// TIA Portal V21 program export: 3 tag tables, 0 data types, 5 data blocks, 7 code blocks (in call order from the OBs), 0 instance data blocks

VAR_GLOBAL   // PLC tag table "DI"
   "DI_PRODUCT SENSOR" AT %I0.0 : Bool;
   "DI_AUTO MANUAL SELECTION" AT %I0.1 : Bool;
   "DI_CYCLE START PB" AT %I0.2 : Bool;
   "DI_CYCLE STOP PB" AT %I0.3 : Bool;
   "DI_EMERGENCY PB" AT %I0.4 : Bool;
   "DI_CONVEYOR VFD FAULT" AT %I0.5 : Bool;
   "DI_SPARE I0.6" AT %I0.6 : Bool;
   "DI_SPARE I0.7" AT %I0.7 : Bool;
   "DI_SPARE I1.0" AT %I1.0 : Bool;
   "DI_SPARE I1.1" AT %I1.1 : Bool;
   "DI_SPARE I1.2" AT %I1.2 : Bool;
   "DI_SPARE I1.3" AT %I1.3 : Bool;
   "DI_SPARE I1.4" AT %I1.4 : Bool;
   "DI_SPARE I1.5" AT %I1.5 : Bool;
END_VAR

VAR_GLOBAL   // PLC tag table "DO"
   "DO_CONVEYOR FWD ON" AT %Q0.0 : Bool;
   "DO_CONVEYOR REV ON" AT %Q0.1 : Bool;
   "DO_FAULT RESET" AT %Q0.2 : Bool;
   "DO_TL GREEN" AT %Q0.3 : Bool;
   "DO_TL RED" AT %Q0.4 : Bool;
   "DO_TL AMBER" AT %Q0.5 : Bool;
   "DO_SPARE Q0.6" AT %Q0.6 : Bool;
   "DO_SPARE Q0.7" AT %Q0.7 : Bool;
   "DO_SPARE Q1.0" AT %Q1.0 : Bool;
   "DO_SPARE Q1.1" AT %Q1.1 : Bool;
END_VAR

VAR_GLOBAL   // PLC tag table "Default tag table"
   System_Byte AT %MB1 : Byte;
   FirstScan AT %M1.0 : Bool;
   DiagStatusUpdate AT %M1.1 : Bool;
   AlwaysTRUE AT %M1.2 : Bool;
   AlwaysFALSE AT %M1.3 : Bool;
   Clock_Byte AT %MB0 : Byte;
   Clock_10Hz AT %M0.0 : Bool;
   Clock_5Hz AT %M0.1 : Bool;
   "Clock_2.5Hz" AT %M0.2 : Bool;
   Clock_2Hz AT %M0.3 : Bool;
   "Clock_1.25Hz" AT %M0.4 : Bool;
   Clock_1Hz AT %M0.5 : Bool;
   "Clock_0.625Hz" AT %M0.6 : Bool;
   "Clock_0.5Hz" AT %M0.7 : Bool;
   "CONTROL ON FLAG" AT %M2.0 : Bool;
   "MANUAL MODE SELECTED" AT %M2.1 : Bool;
   "AUTO MODE SELECTED" AT %M2.2 : Bool;
   "FAULT RESET FLAG" AT %M2.3 : Bool;
   "FAULT BIT" AT %M2.4 : Bool;
   "MANUAL CONVEYOR FWD ON FLAG" AT %M2.5 : Bool;
   "MANUAL CONVEYOR REV ON FLAG" AT %M2.6 : Bool;
END_VAR

DATA_BLOCK "DB_ALARMS"   // DB2
{ S7_Optimized_Access := 'FALSE' }
VERSION : 0.1
// stored: AutoNumber true, DBAccessibleFromOPCUA true, IsOnlyStoredInLoadMemory false, IsWriteProtectedInAS false
   VAR
      "EMERGENCY PB PRESSED FAULT" : Bool;
      "VFD FAULT" : Bool;
      SPARE1 : Bool;
      SPARE2 : Bool;
      SPARE3 : Bool;
      SPARE4 : Bool;
      SPARE5 : Bool;
      SPARE6 : Bool;
      SPARE7 : Bool;
      SPARE8 : Bool;
      SPARE9 : Bool;
      SPARE10 : Bool;
      SPARE11 : Bool;
      SPARE12 : Bool;
      SPARE13 : Bool;
      SPARE14 : Bool;
      "FAULT POP" : Bool;
      "WARNING POP" : Bool;
   END_VAR
BEGIN
END_DATA_BLOCK

DATA_BLOCK "DB_AUTO"   // DB3
{ S7_Optimized_Access := 'FALSE' }
VERSION : 0.1
// stored: AutoNumber true, DBAccessibleFromOPCUA true, IsOnlyStoredInLoadMemory false, IsWriteProtectedInAS false
   VAR
      ACTIVE : Bool;
      "CONVEYOR ON" : Bool;
      "CONVEYOR OFF1" : Bool;
      "CONVEYOR OFF2" : Bool;
      P_TRG : Bool;
      "CAMERA DONE" : Bool;
      "AUTO STATUS" : Int;
      "STOP DELAY TIMER" : IEC_TIMER;
      "SENSOR CHECK DELAY" { S7_SetPoint := 'True'} : IEC_TIMER;
   END_VAR
BEGIN
END_DATA_BLOCK

DATA_BLOCK "DB_CAMERA"   // DB5
{ S7_Optimized_Access := 'FALSE' }
VERSION : 0.1
// stored: AutoNumber true, DBAccessibleFromOPCUA true, IsOnlyStoredInLoadMemory false, IsWriteProtectedInAS false
   VAR
      DATA1 : Int;
      DATA2 : Int;
      DATA3 : Int;
      DATA4 : Int;
      DATA5 : Int;
      DATA6 : Int;
      DATA7 : Int;
      DATA8 : Int;
      DATA9 : Int;
      DATA10 : Int;
      DATA11 : Int;
      DATA12 : Int;
      DATA13 : Int;
      DATA14 : Int;
      DATA15 : Int;
      DATA16 : Int;
      DATA17 : Int;
      DATA18 : Int;
      DATA19 : Int;
   END_VAR
BEGIN
END_DATA_BLOCK

DATA_BLOCK "DB_HMI"   // DB1
{ S7_Optimized_Access := 'FALSE' }
VERSION : 0.1
// stored: AutoNumber true, DBAccessibleFromOPCUA true, IsOnlyStoredInLoadMemory false, IsWriteProtectedInAS false
   VAR RETAIN
      "FAULT RESET PB" : Bool;
      "MOTOR JOG FWD PB" : Bool;
      "MOTOR JOG REV PB" : Bool;
      "STOP TIME" : DInt;
      "CAMERA DONE" : Bool;
   END_VAR
BEGIN
END_DATA_BLOCK

DATA_BLOCK "DB_TCP_IP"   // DB12
{ S7_Optimized_Access := 'TRUE' }
VERSION : 0.1
// stored: AutoNumber true, DBAccessibleFromOPCUA true, IsOnlyStoredInLoadMemory false, IsRetainMemResEnabled false, IsWriteProtectedInAS false, MemoryReserve 100
   VAR
      "MY CONNECT DATA" { S7_SetPoint := 'True'} : TCON_IP_v4;
      "NO OF DONE" { S7_SetPoint := 'True'} : UDInt;
      "NO OF ERROR" : UDInt;
      "ERROR STATUS" : UDInt;
   END_VAR
BEGIN
END_DATA_BLOCK

ORGANIZATION_BLOCK "Main"   // OB1, LAD, ProgramCycle
TITLE = "Main Program Sweep (Cycle)"
{ S7_Optimized_Access := 'TRUE' }
VERSION : 0.1
// stored: AutoNumber true, IsIECCheckEnabled false, SetENOAutomatically false
   VAR_INPUT
      Initial_Call : Bool;   // Initial call of this OB
      Remanence : Bool;   // =True, if remanent data are available
   END_VAR
BEGIN

REGION Network 1
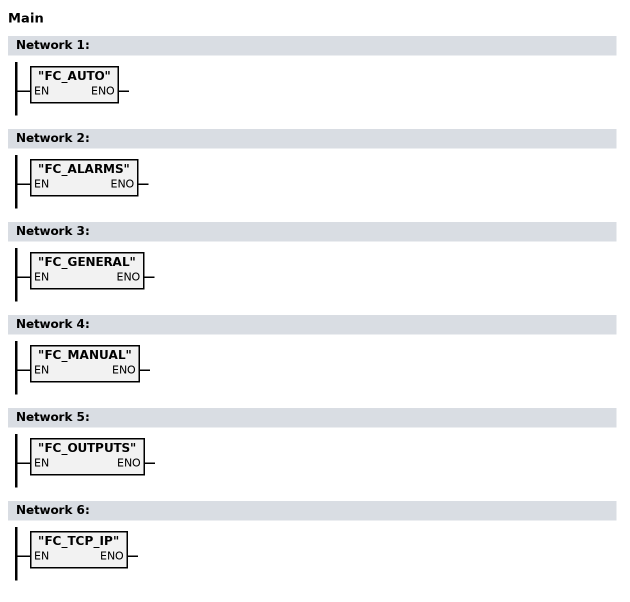
   RUNG wire#powerrail
      "FC_AUTO"()
   END_RUNG
   // the same network as SCL:
   "FC_AUTO"();
END_REGION

REGION Network 2
   RUNG wire#powerrail
      "FC_ALARMS"()
   END_RUNG
   // the same network as SCL:
   "FC_ALARMS"();
END_REGION

REGION Network 3
   RUNG wire#powerrail
      "FC_GENERAL"()
   END_RUNG
   // the same network as SCL:
   "FC_GENERAL"();
END_REGION

REGION Network 4
   RUNG wire#powerrail
      "FC_MANUAL"()
   END_RUNG
   // the same network as SCL:
   "FC_MANUAL"();
END_REGION

REGION Network 5
   RUNG wire#powerrail
      "FC_OUTPUTS"()
   END_RUNG
   // the same network as SCL:
   "FC_OUTPUTS"();
END_REGION

REGION Network 6
   RUNG wire#powerrail
      "FC_TCP_IP"()
   END_RUNG
   // the same network as SCL:
   "FC_TCP_IP"();
END_REGION
END_ORGANIZATION_BLOCK

FUNCTION "FC_AUTO" : Void   // FC5, LAD
{ S7_Optimized_Access := 'TRUE' }
VERSION : 0.1
// stored: AutoNumber true, IsIECCheckEnabled false, SetENOAutomatically false, UDAEnableTagReadback false
   VAR_TEMP   // added for the SCL form of the ladder/FBD networks
      _w1 : Bool;
      _w2 : Bool;
      _w3 : Bool;
   END_VAR
BEGIN

REGION Network 1: AUTO ON
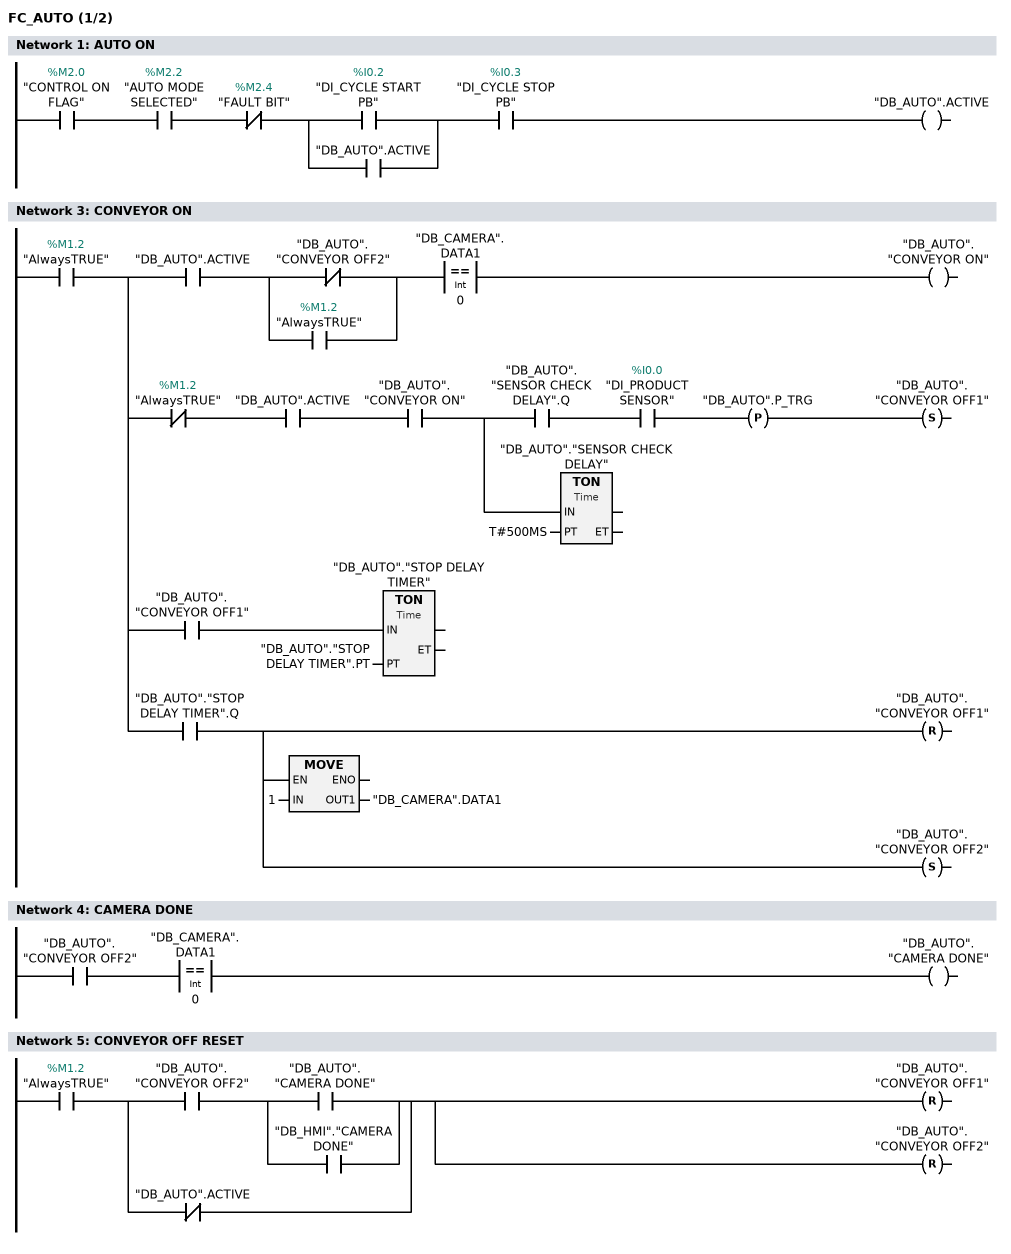
   RUNG wire#powerrail
      Contact( "CONTROL ON FLAG" )
      Contact( "AUTO MODE SELECTED" )
      I_Contact( "FAULT BIT" )
      wire#w1
      Contact( "DI_CYCLE START PB" )
      wire#w2
      Contact( "DI_CYCLE STOP PB" )
      Coil( "DB_AUTO".ACTIVE )
   END_RUNG
   RUNG wire#w1
      Contact( "DB_AUTO".ACTIVE )
   END_RUNG wire#w2
   // the same network as SCL:
   "DB_AUTO".ACTIVE := "CONTROL ON FLAG" AND "AUTO MODE SELECTED" AND NOT "FAULT BIT" AND ("DI_CYCLE START PB" OR "DB_AUTO".ACTIVE) AND "DI_CYCLE STOP PB";
END_REGION

REGION Network 2 (SCL): STOP DELAY TIME
   "DB_AUTO"."STOP DELAY TIMER".PT := "DB_HMI"."STOP TIME" * 1000;
END_REGION

REGION Network 3: CONVEYOR ON
   RUNG wire#powerrail
      Contact( "AlwaysTRUE" )
      wire#w1
      Contact( "DB_AUTO".ACTIVE )
      wire#w2
      I_Contact( "DB_AUTO"."CONVEYOR OFF2" )
      wire#w3
      { S7_Templates := "SrcType := Int" } EQ_Contact(in1 := "DB_CAMERA".DATA1, in2 := 0)
      Coil( "DB_AUTO"."CONVEYOR ON" )
   END_RUNG
   RUNG wire#w2
      Contact( "AlwaysTRUE" )
   END_RUNG wire#w3
   RUNG wire#w1
      I_Contact( "AlwaysTRUE" )
      Contact( "DB_AUTO".ACTIVE )
      Contact( "DB_AUTO"."CONVEYOR ON" )
      wire#w4
      Contact( "DB_AUTO"."SENSOR CHECK DELAY".Q )
      Contact( "DI_PRODUCT SENSOR" )
      P_Trig( "DB_AUTO".P_TRG )
      S_Coil( "DB_AUTO"."CONVEYOR OFF1" )
   END_RUNG
   RUNG wire#w4
      { S7_Templates := "time_type := Time" } "DB_AUTO"."SENSOR CHECK DELAY".TON(pt := T#500MS, et =>)
   END_RUNG
   RUNG wire#w1
      Contact( "DB_AUTO"."CONVEYOR OFF1" )
      { S7_Templates := "time_type := Time" } "DB_AUTO"."STOP DELAY TIMER".TON(pt := "DB_AUTO"."STOP DELAY TIMER".PT, et =>)
   END_RUNG
   RUNG wire#w1
      Contact( "DB_AUTO"."STOP DELAY TIMER".Q )
      wire#w5
      R_Coil( "DB_AUTO"."CONVEYOR OFF1" )
   END_RUNG
   RUNG wire#w5
      Move(in := 1, out1 => "DB_CAMERA".DATA1)
   END_RUNG
   RUNG wire#w5
      S_Coil( "DB_AUTO"."CONVEYOR OFF2" )
   END_RUNG
   // the same network as SCL:
   "DB_AUTO"."CONVEYOR ON" := "AlwaysTRUE" AND "DB_AUTO".ACTIVE AND (NOT "DB_AUTO"."CONVEYOR OFF2" OR "AlwaysTRUE") AND ("DB_CAMERA".DATA1 = 0);
   #_w1 := "AlwaysTRUE" AND NOT "AlwaysTRUE" AND "DB_AUTO".ACTIVE AND "DB_AUTO"."CONVEYOR ON";
   #_w2 := #_w1 AND "DB_AUTO"."SENSOR CHECK DELAY".Q AND "DI_PRODUCT SENSOR";
   #_w3 := #_w2 AND NOT "DB_AUTO".P_TRG;   // rising edge
   "DB_AUTO".P_TRG := #_w2;
   IF #_w3 THEN "DB_AUTO"."CONVEYOR OFF1" := TRUE; END_IF;
   "DB_AUTO"."SENSOR CHECK DELAY".TON(IN := #_w1, PT := T#500MS);
   "DB_AUTO"."STOP DELAY TIMER".TON(IN := "AlwaysTRUE" AND "DB_AUTO"."CONVEYOR OFF1",
                           PT := "DB_AUTO"."STOP DELAY TIMER".PT);
   IF "AlwaysTRUE" AND "DB_AUTO"."STOP DELAY TIMER".Q THEN
       "DB_AUTO"."CONVEYOR OFF1" := FALSE;
       "DB_CAMERA".DATA1 := 1;
       "DB_AUTO"."CONVEYOR OFF2" := TRUE;
   END_IF;
END_REGION

REGION Network 4: CAMERA DONE
   RUNG wire#powerrail
      Contact( "DB_AUTO"."CONVEYOR OFF2" )
      { S7_Templates := "SrcType := Int" } EQ_Contact(in1 := "DB_CAMERA".DATA1, in2 := 0)
      Coil( "DB_AUTO"."CAMERA DONE" )
   END_RUNG
   // the same network as SCL:
   "DB_AUTO"."CAMERA DONE" := "DB_AUTO"."CONVEYOR OFF2" AND ("DB_CAMERA".DATA1 = 0);
END_REGION

REGION Network 5: CONVEYOR OFF RESET
   RUNG wire#powerrail
      Contact( "AlwaysTRUE" )
      wire#w1
      Contact( "DB_AUTO"."CONVEYOR OFF2" )
      wire#w2
      Contact( "DB_AUTO"."CAMERA DONE" )
      wire#w3
      R_Coil( "DB_AUTO"."CONVEYOR OFF1" )
   END_RUNG
   RUNG wire#w2
      Contact( "DB_HMI"."CAMERA DONE" )
   END_RUNG wire#w3
   RUNG wire#w1
      I_Contact( "DB_AUTO".ACTIVE )
   END_RUNG wire#w3
   RUNG wire#w3
      R_Coil( "DB_AUTO"."CONVEYOR OFF2" )
   END_RUNG
   // the same network as SCL:
   IF "AlwaysTRUE" AND (("DB_AUTO"."CONVEYOR OFF2" AND ("DB_AUTO"."CAMERA DONE" OR "DB_HMI"."CAMERA DONE")) OR NOT "DB_AUTO".ACTIVE) THEN
       "DB_AUTO"."CONVEYOR OFF1" := FALSE;
       "DB_AUTO"."CONVEYOR OFF2" := FALSE;
   END_IF;
END_REGION

REGION Network 6: AUTO STATUS
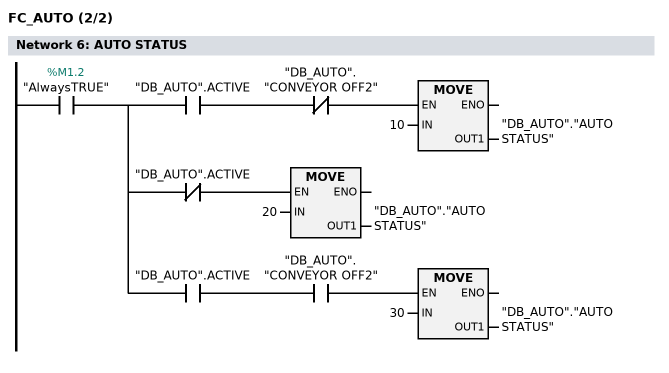
   RUNG wire#powerrail
      Contact( "AlwaysTRUE" )
      wire#w1
      Contact( "DB_AUTO".ACTIVE )
      I_Contact( "DB_AUTO"."CONVEYOR OFF2" )
      Move(in := 10, out1 => "DB_AUTO"."AUTO STATUS")
   END_RUNG
   RUNG wire#w1
      I_Contact( "DB_AUTO".ACTIVE )
      Move(in := 20, out1 => "DB_AUTO"."AUTO STATUS")
   END_RUNG
   RUNG wire#w1
      Contact( "DB_AUTO".ACTIVE )
      Contact( "DB_AUTO"."CONVEYOR OFF2" )
      Move(in := 30, out1 => "DB_AUTO"."AUTO STATUS")
   END_RUNG
   // the same network as SCL:
   IF "AlwaysTRUE" AND "DB_AUTO".ACTIVE AND NOT "DB_AUTO"."CONVEYOR OFF2" THEN
       "DB_AUTO"."AUTO STATUS" := 10;
   END_IF;
   IF "AlwaysTRUE" AND NOT "DB_AUTO".ACTIVE THEN "DB_AUTO"."AUTO STATUS" := 20; END_IF;
   IF "AlwaysTRUE" AND "DB_AUTO".ACTIVE AND "DB_AUTO"."CONVEYOR OFF2" THEN
       "DB_AUTO"."AUTO STATUS" := 30;
   END_IF;
END_REGION
END_FUNCTION

FUNCTION "FC_ALARMS" : Void   // FC3, LAD
{ S7_Optimized_Access := 'TRUE' }
VERSION : 0.1
// stored: AutoNumber true, IsIECCheckEnabled false, SetENOAutomatically false, UDAEnableTagReadback false
BEGIN

REGION Network 1: EMERGENCY PB PRESSED FAULT (I0.4)
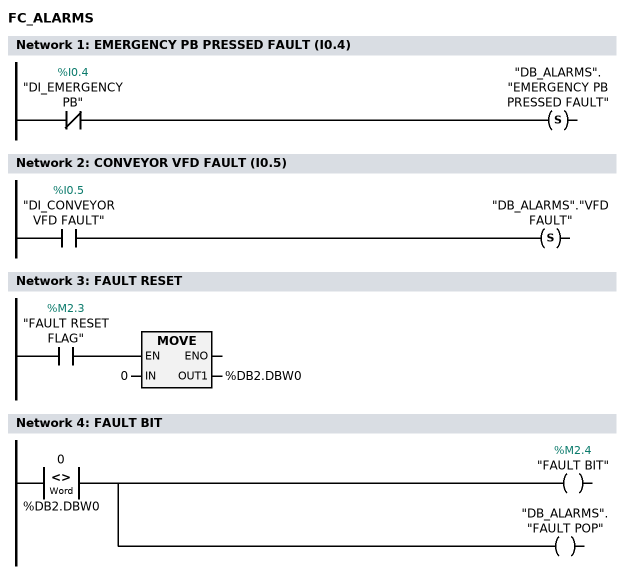
   RUNG wire#powerrail
      I_Contact( "DI_EMERGENCY PB" )
      S_Coil( "DB_ALARMS"."EMERGENCY PB PRESSED FAULT" )
   END_RUNG
   // the same network as SCL:
   IF NOT "DI_EMERGENCY PB" THEN "DB_ALARMS"."EMERGENCY PB PRESSED FAULT" := TRUE; END_IF;
END_REGION

REGION Network 2: CONVEYOR VFD FAULT (I0.5)
   RUNG wire#powerrail
      Contact( "DI_CONVEYOR VFD FAULT" )
      S_Coil( "DB_ALARMS"."VFD FAULT" )
   END_RUNG
   // the same network as SCL:
   IF "DI_CONVEYOR VFD FAULT" THEN "DB_ALARMS"."VFD FAULT" := TRUE; END_IF;
END_REGION

REGION Network 3: FAULT RESET
   RUNG wire#powerrail
      Contact( "FAULT RESET FLAG" )
      Move(in := 0, out1 => %DB2.DBW0)
   END_RUNG
   // the same network as SCL:
   IF "FAULT RESET FLAG" THEN %DB2.DBW0 := 0; END_IF;
END_REGION

REGION Network 4: FAULT BIT
   RUNG wire#powerrail
      { S7_Templates := "SrcType := Word" } NE_Contact(in1 := 0, in2 := %DB2.DBW0)
      wire#w1
      Coil( "FAULT BIT" )
   END_RUNG
   RUNG wire#w1
      Coil( "DB_ALARMS"."FAULT POP" )
   END_RUNG
   // the same network as SCL:
   "FAULT BIT" := 0 <> %DB2.DBW0;
   "DB_ALARMS"."FAULT POP" := "FAULT BIT";
END_REGION
END_FUNCTION

FUNCTION "FC_GENERAL" : Void   // FC1, LAD
{ S7_Optimized_Access := 'TRUE' }
VERSION : 0.1
// stored: AutoNumber true, IsIECCheckEnabled false, SetENOAutomatically false, UDAEnableTagReadback false
BEGIN

REGION Network 1: CONTROL ON
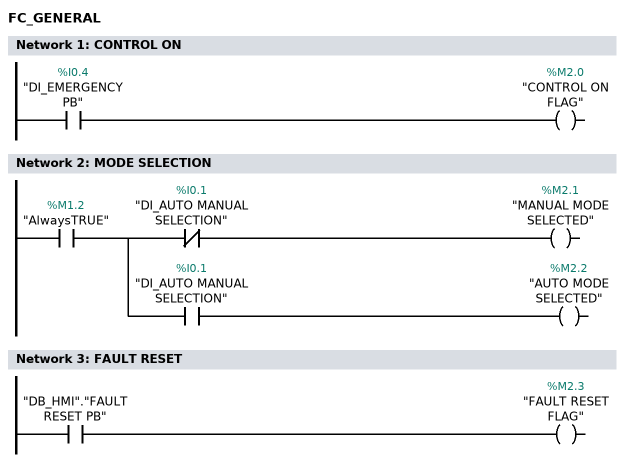
   RUNG wire#powerrail
      Contact( "DI_EMERGENCY PB" )
      Coil( "CONTROL ON FLAG" )
   END_RUNG
   // the same network as SCL:
   "CONTROL ON FLAG" := "DI_EMERGENCY PB";
END_REGION

REGION Network 2: MODE SELECTION
   RUNG wire#powerrail
      Contact( "AlwaysTRUE" )
      wire#w1
      I_Contact( "DI_AUTO MANUAL SELECTION" )
      Coil( "MANUAL MODE SELECTED" )
   END_RUNG
   RUNG wire#w1
      Contact( "DI_AUTO MANUAL SELECTION" )
      Coil( "AUTO MODE SELECTED" )
   END_RUNG
   // the same network as SCL:
   "MANUAL MODE SELECTED" := "AlwaysTRUE" AND NOT "DI_AUTO MANUAL SELECTION";
   "AUTO MODE SELECTED" := "AlwaysTRUE" AND "DI_AUTO MANUAL SELECTION";
END_REGION

REGION Network 3: FAULT RESET
   RUNG wire#powerrail
      Contact( "DB_HMI"."FAULT RESET PB" )
      Coil( "FAULT RESET FLAG" )
   END_RUNG
   // the same network as SCL:
   "FAULT RESET FLAG" := "DB_HMI"."FAULT RESET PB";
END_REGION
END_FUNCTION

FUNCTION "FC_MANUAL" : Void   // FC2, LAD
{ S7_Optimized_Access := 'TRUE' }
VERSION : 0.1
// stored: AutoNumber true, IsIECCheckEnabled false, SetENOAutomatically false, UDAEnableTagReadback false
   VAR_TEMP   // added for the SCL form of the ladder/FBD networks
      _w1 : Bool;
   END_VAR
BEGIN

REGION Network 1: MOTOR FWD /REV ON
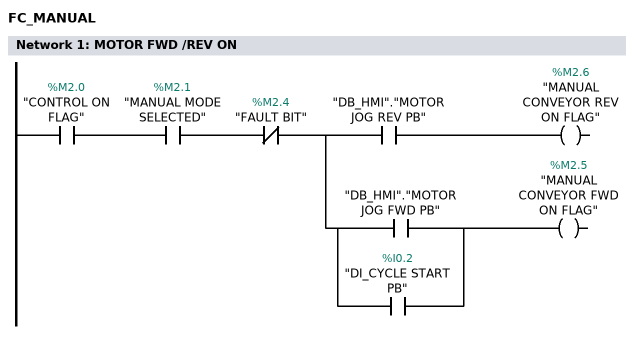
   RUNG wire#powerrail
      Contact( "CONTROL ON FLAG" )
      Contact( "MANUAL MODE SELECTED" )
      I_Contact( "FAULT BIT" )
      wire#w1
      Contact( "DB_HMI"."MOTOR JOG REV PB" )
      Coil( "MANUAL CONVEYOR REV ON FLAG" )
   END_RUNG
   RUNG wire#w1
      Contact( "DB_HMI"."MOTOR JOG FWD PB" )
      wire#w2
      Coil( "MANUAL CONVEYOR FWD ON FLAG" )
   END_RUNG
   RUNG wire#w1
      Contact( "DI_CYCLE START PB" )
   END_RUNG wire#w2
   // the same network as SCL:
   #_w1 := "CONTROL ON FLAG" AND "MANUAL MODE SELECTED" AND NOT "FAULT BIT";
   "MANUAL CONVEYOR REV ON FLAG" := #_w1 AND "DB_HMI"."MOTOR JOG REV PB";
   "MANUAL CONVEYOR FWD ON FLAG" := #_w1 AND ("DB_HMI"."MOTOR JOG FWD PB" OR "DI_CYCLE START PB");
END_REGION
END_FUNCTION

FUNCTION "FC_OUTPUTS" : Void   // FC4, LAD
{ S7_Optimized_Access := 'TRUE' }
VERSION : 0.1
// stored: AutoNumber true, IsIECCheckEnabled false, SetENOAutomatically false, UDAEnableTagReadback false
BEGIN

REGION Network 1: CONVEYOR FWD ON
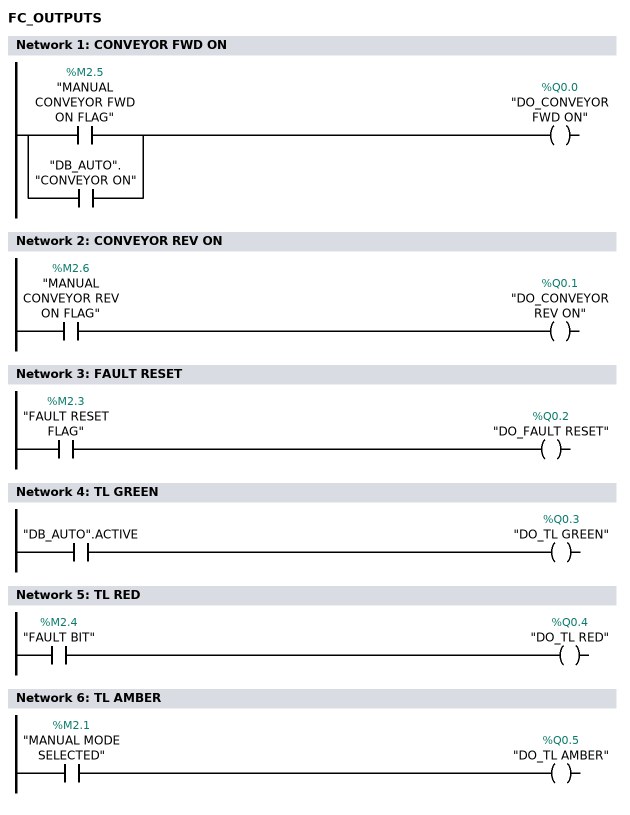
   RUNG wire#powerrail
      Contact( "MANUAL CONVEYOR FWD ON FLAG" )
      wire#w1
      Coil( "DO_CONVEYOR FWD ON" )
   END_RUNG
   RUNG wire#powerrail
      Contact( "DB_AUTO"."CONVEYOR ON" )
   END_RUNG wire#w1
   // the same network as SCL:
   "DO_CONVEYOR FWD ON" := "MANUAL CONVEYOR FWD ON FLAG" OR "DB_AUTO"."CONVEYOR ON";
END_REGION

REGION Network 2: CONVEYOR REV ON
   RUNG wire#powerrail
      Contact( "MANUAL CONVEYOR REV ON FLAG" )
      Coil( "DO_CONVEYOR REV ON" )
   END_RUNG
   // the same network as SCL:
   "DO_CONVEYOR REV ON" := "MANUAL CONVEYOR REV ON FLAG";
END_REGION

REGION Network 3: FAULT RESET
   RUNG wire#powerrail
      Contact( "FAULT RESET FLAG" )
      Coil( "DO_FAULT RESET" )
   END_RUNG
   // the same network as SCL:
   "DO_FAULT RESET" := "FAULT RESET FLAG";
END_REGION

REGION Network 4: TL GREEN
   RUNG wire#powerrail
      Contact( "DB_AUTO".ACTIVE )
      Coil( "DO_TL GREEN" )
   END_RUNG
   // the same network as SCL:
   "DO_TL GREEN" := "DB_AUTO".ACTIVE;
END_REGION

REGION Network 5: TL RED
   RUNG wire#powerrail
      Contact( "FAULT BIT" )
      Coil( "DO_TL RED" )
   END_RUNG
   // the same network as SCL:
   "DO_TL RED" := "FAULT BIT";
END_REGION

REGION Network 6: TL AMBER
   RUNG wire#powerrail
      Contact( "MANUAL MODE SELECTED" )
      Coil( "DO_TL AMBER" )
   END_RUNG
   // the same network as SCL:
   "DO_TL AMBER" := "MANUAL MODE SELECTED";
END_REGION
END_FUNCTION

FUNCTION "FC_TCP_IP" : Void   // FC6, LAD
{ S7_Optimized_Access := 'TRUE' }
VERSION : 0.1
// stored: AutoNumber true, IsIECCheckEnabled false, SetENOAutomatically false, UDAEnableTagReadback false
BEGIN

REGION Network 1: Connection definition
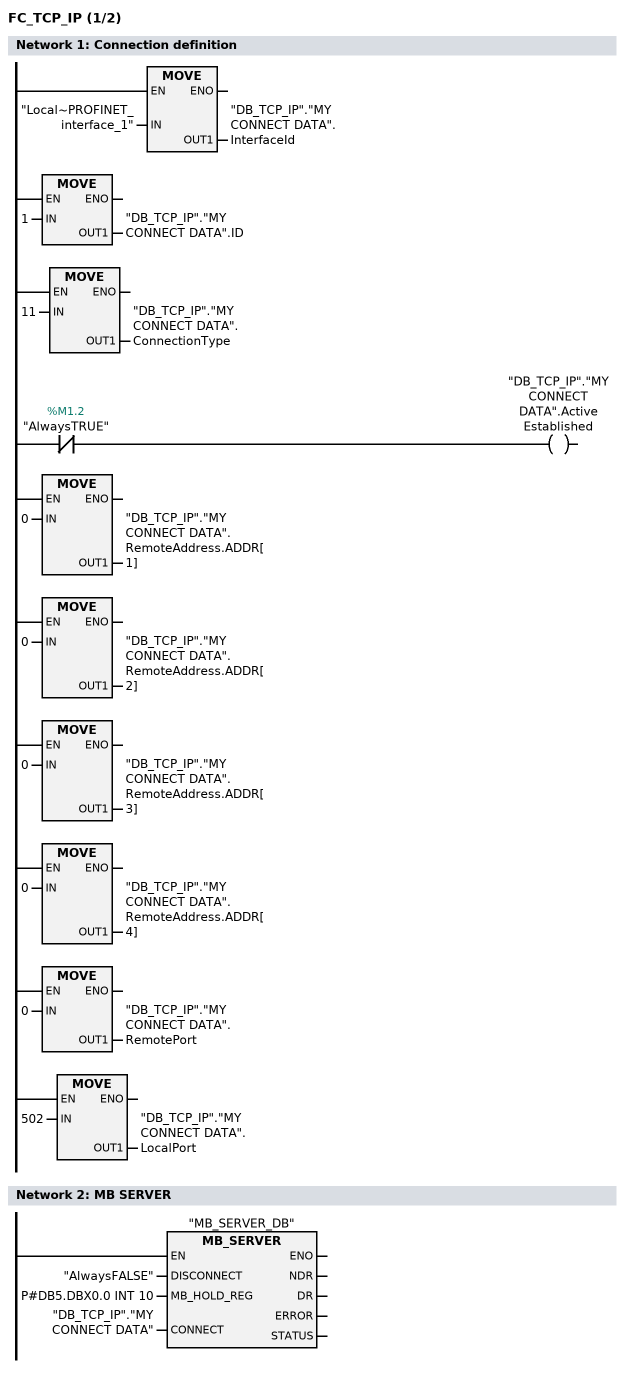
   RUNG wire#powerrail
      Move(in := "Local~PROFINET_interface_1", out1 => "DB_TCP_IP"."MY CONNECT DATA".InterfaceId)
   END_RUNG
   RUNG wire#powerrail
      Move(in := 1, out1 => "DB_TCP_IP"."MY CONNECT DATA".ID)
   END_RUNG
   RUNG wire#powerrail
      Move(in := 11, out1 => "DB_TCP_IP"."MY CONNECT DATA".ConnectionType)
   END_RUNG
   RUNG wire#powerrail
      I_Contact( "AlwaysTRUE" )
      Coil( "DB_TCP_IP"."MY CONNECT DATA".ActiveEstablished )
   END_RUNG
   RUNG wire#powerrail
      Move(in := 0, out1 => "DB_TCP_IP"."MY CONNECT DATA".RemoteAddress.ADDR[1])
   END_RUNG
   RUNG wire#powerrail
      Move(in := 0, out1 => "DB_TCP_IP"."MY CONNECT DATA".RemoteAddress.ADDR[2])
   END_RUNG
   RUNG wire#powerrail
      Move(in := 0, out1 => "DB_TCP_IP"."MY CONNECT DATA".RemoteAddress.ADDR[3])
   END_RUNG
   RUNG wire#powerrail
      Move(in := 0, out1 => "DB_TCP_IP"."MY CONNECT DATA".RemoteAddress.ADDR[4])
   END_RUNG
   RUNG wire#powerrail
      Move(in := 0, out1 => "DB_TCP_IP"."MY CONNECT DATA".RemotePort)
   END_RUNG
   RUNG wire#powerrail
      Move(in := 502, out1 => "DB_TCP_IP"."MY CONNECT DATA".LocalPort)
   END_RUNG
   // the same network as SCL:
   "DB_TCP_IP"."MY CONNECT DATA".InterfaceId := "Local~PROFINET_interface_1";
   "DB_TCP_IP"."MY CONNECT DATA".ID := 1;
   "DB_TCP_IP"."MY CONNECT DATA".ConnectionType := 11;
   "DB_TCP_IP"."MY CONNECT DATA".ActiveEstablished := NOT "AlwaysTRUE";
   "DB_TCP_IP"."MY CONNECT DATA".RemoteAddress.ADDR[1] := 0;
   "DB_TCP_IP"."MY CONNECT DATA".RemoteAddress.ADDR[2] := 0;
   "DB_TCP_IP"."MY CONNECT DATA".RemoteAddress.ADDR[3] := 0;
   "DB_TCP_IP"."MY CONNECT DATA".RemoteAddress.ADDR[4] := 0;
   "DB_TCP_IP"."MY CONNECT DATA".RemotePort := 0;
   "DB_TCP_IP"."MY CONNECT DATA".LocalPort := 502;
END_REGION

REGION Network 2: MB SERVER
   RUNG wire#powerrail
      "MB_SERVER_DB".MB_SERVER(DISCONNECT := "AlwaysFALSE", MB_HOLD_REG := P#DB5.DBX0.0 INT 10, CONNECT := "DB_TCP_IP"."MY CONNECT DATA", NDR =>, DR =>, ERROR =>, STATUS =>)
   END_RUNG
   // the same network as SCL:
   "MB_SERVER_DB"(DISCONNECT := "AlwaysFALSE",   // MB_SERVER
                  MB_HOLD_REG := P#DB5.DBX0.0 INT 10,
                  CONNECT := "DB_TCP_IP"."MY CONNECT DATA");
END_REGION

REGION Network 3: ERROR CHECK
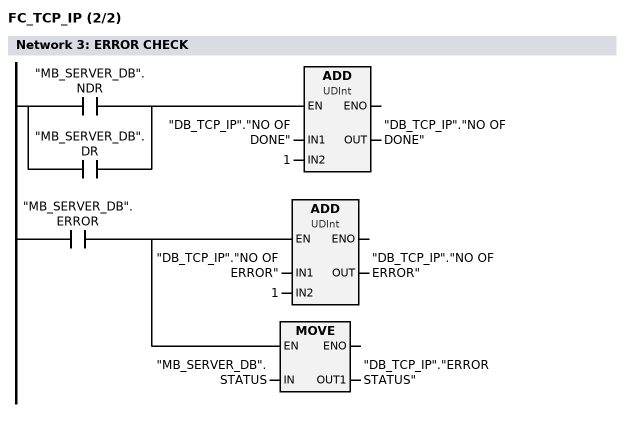
   RUNG wire#powerrail
      Contact( "MB_SERVER_DB".NDR )
      wire#w1
      { S7_Templates := "SrcType := UDInt" } Add(in1 := "DB_TCP_IP"."NO OF DONE", in2 := 1, out => "DB_TCP_IP"."NO OF DONE")
   END_RUNG
   RUNG wire#powerrail
      Contact( "MB_SERVER_DB".DR )
   END_RUNG wire#w1
   RUNG wire#powerrail
      Contact( "MB_SERVER_DB".ERROR )
      wire#w2
      { S7_Templates := "SrcType := UDInt" } Add(in1 := "DB_TCP_IP"."NO OF ERROR", in2 := 1, out => "DB_TCP_IP"."NO OF ERROR")
   END_RUNG
   RUNG wire#w2
      Move(in := "MB_SERVER_DB".STATUS, out1 => "DB_TCP_IP"."ERROR STATUS")
   END_RUNG
   // the same network as SCL:
   IF "MB_SERVER_DB".NDR OR "MB_SERVER_DB".DR THEN
       "DB_TCP_IP"."NO OF DONE" := "DB_TCP_IP"."NO OF DONE" + 1;
   END_IF;
   IF "MB_SERVER_DB".ERROR THEN
       "DB_TCP_IP"."NO OF ERROR" := "DB_TCP_IP"."NO OF ERROR" + 1;
       "DB_TCP_IP"."ERROR STATUS" := "MB_SERVER_DB".STATUS;
   END_IF;
END_REGION
END_FUNCTION
